Fanuc KAREL source: KO00115.KL

PROGRAM KO00115
%NOLOCKGROUP
VAR
  A: ARRAY[2] OF BYTE
  B: REAL
  OUT: INTEGER
BEGIN
  A[1] = 1
  B = 2
  OUT = ATAN2(A[1], B)
END KO00115
